Staubli VAL3: initLabel.pgx

public program initLabel(utLabel& x_utLabel[], string x_sPage, string x_sId, string x_sText)
begin
  x_utLabel.Common.sPage=x_sPage
  x_utLabel.Common.sID=x_sId
  userPageBind(x_utLabel.Common.sPage,x_utLabel.Common.sID,"innerHTML",x_utLabel.Common.sText,1,"r")
  //userPageBind(x_sPage,x_utLabel.Common.sID,"style.backgroundColor",x_utLabel.Appearance.sBackgroundColour,1,"r")
  //userPageBindClick(x_sPage,x_utLabel.Common.sID,x_utLabel.Events.bClick,true)
  //
  if x_sText=="" or x_sText=="Null"
    x_utLabel.Common.sText=""
  else
    x_utLabel.Common.sText=x_sText
  endIf
  //x_utLabel.Appearance.sBackgroundColour="#F3F4F4"
  x_utLabel.Data.nVal=99
end
